Yaskawa INFORM job: CA.JBI

/JOB
//NAME CA
//POS
///NPOS 12,0,0,0,0,0
///TOOL 0
///POSTYPE PULSE
///PULSE
C00000=1,-60004,-60001,1,-90000,0
C00001=-1984,15242,-61866,-97156,-4498,46014
C00002=-2791,22019,-61532,-135569,-7364,64330
C00003=-4032,20706,-63624,-134675,-7979,64252
C00004=-5437,22381,-61136,-129323,-7982,62109
C00005=-5232,23076,-55377,-106480,-6075,51263
C00006=-5865,26630,-54490,-120600,-7233,58100
C00007=-2562,24508,-57771,-132424,-6780,62782
C00008=-6115,23060,-59812,-125768,-7891,60614
C00009=-4384,24352,-57852,-127531,-7192,60971
C00010=-4384,19661,-55926,-86417,-5382,41587
C00011=1,-60004,-60001,1,-90000,0
//INST
///DATE 2026/06/19 13:02
///ATTR SC,RW
///GROUP1 RB1
NOP
MOVJ C00000 VJ=0.73
MOVJ C00001 VJ=15.00
MOVC C00002 V=11.0
ARCON ASF#(13)
MOVC C00003 V=11.0
MOVC C00004 V=11.0
ARCOF AEF#(13)
MOVL C00005 V=11.0
MOVL C00006 V=11.0
ARCON ASF#(13)
MOVL C00007 V=11.0
MOVL C00008 V=11.0
ARCOF AEF#(13)
MOVL C00009 V=11.0
ARCON ASF#(13)
TIMER T=0.50
ARCOF AEF#(13)
MOVL C00010 V=11.0
MOVJ C00011 VJ=15.00
END
